DATA_BLOCK "LineData"
{ S7_Optimized_Access := 'TRUE' }
VERSION : 0.1
NON_RETAIN
"FillingLine"

BEGIN

END_DATA_BLOCK

